Fanuc KAREL source: kt00533.KL

PROGRAM KT00533
%STACKSIZE=65535
%PRIORITY=65535
%NOLOCKGROUP
VAR
P1 : JOINTPOS9
P2 : POSITION
OUT : BOOLEAN
BEGIN
-- UNRESOLVED_PC line 8 opcodes [49 7E 49 AC 23] marker_code=0
END KT00533
